{attribute 'TcGvlVarFlags' := 'OPC'}
VAR_GLOBAL
    // EL3702 analog input data — written by FB_AnalogInHandler, read by Python over ADS
    // ADS symbol: GVL_AnalogIn.stAnalogIn
    stAnalogIn1         : ST_AnalogInData;
    stAnalogIn2         : ST_AnalogInData;
END_VAR

(* stored: Version 1.1.0.1, ProductVersion 3.1.4026.18
   GVL GVL_AnalogIn: Id {41d41d25-dcb4-4550-97a6-bccb4f741935} *)
